(*
SPDX-FileCopyrightText: © 2026 Oleksandr Tiutyk <trofimich@gmail.com>
SPDX-License-Identifier: MIT
License: https://opensource.org/license/mit
*)

(*!
<summary>Enumerates allocated text fragments from a borrowed source string.</summary>
<description>
Initialization requires a separator containing 1 to 80 characters, stored in a fixed buffer. The source must
remain alive and unchanged during iteration. The enumerator owns the current fragment; borrowed fragment
references expire on MoveNext, Reset or destruction. Allocation failure uses the terminal memory mechanism.
With a nonempty separator, empty fragments are preserved when RemoveEmptyEntries is FALSE, including the final
fragment after a trailing separator and one fragment for an empty source. RemoveEmptyEntries filters empty
fragments after optional trimming. MaxCount still limits the number of returned fragments. Do not copy an
instance by assignment or pass it by value while it owns an allocated buffer; use references instead.
Assignment does not clone the buffer or transfer ownership. Do not overwrite an instance that still owns a
buffer. The creator is responsible for the splitter lifetime and cleanup. Release the current fragment with
Reset when abandoning iteration. Delete the splitter itself only if it was allocated with __NEW; FB_exit
releases its current fragment. Statically or locally declared instances must not be passed to __DELETE. The
borrowed source is never owned or freed by the splitter.
</description>
*)

{attribute 'no_explicit_call' := 'do not call this function block directly'}
FUNCTION_BLOCK WideStringSplittingEnumerator EXTENDS Object IMPLEMENTS IEnumerator
VAR_OUTPUT
	SourceString : POINTER TO WSTRING;
	SourceStringLength : UDINT;
	SourceStringSize : UDINT;
	Separator : WSTRING(80);
	SeparatorLength : UDINT;
	//!<summary>
	//! Maximum number of returned fragments; zero means unlimited. Empty fragments removed after optional
	//! trimming do not count toward the limit. Remaining text is not returned after the limit is reached and is
	//! not merged into the last fragment.
	//! </summary>
	MaxCount : UDINT := 0;
	TrimEntries : BOOL := FALSE;
	RemoveEmptyEntries : BOOL := FALSE;	
END_VAR
VAR_STAT
	//! <summary>Class name shared by all instances of this function block.</summary>
	{attribute 'hide'} 
	_ClassName : STRING := __POUNAME();
END_VAR
VAR
	{attribute 'hide'} 
	_CurrentString : POINTER TO WSTRING;
	{attribute 'hide'} 
	_CurrentStringLength : UDINT;
	{attribute 'hide'} 
	_CurrentEntry : POINTER TO WSTRING;
	{attribute 'hide'} 
	_CurrentEntrySize : UDINT;
	{attribute 'hide'} 
	_EntryCount : UDINT; 
END_VAR

{attribute 'monitoring' := 'call'}
PROPERTY ClassName : REFERENCE TO STRING
GET
ClassName REF= _ClassName;
END_GET
END_PROPERTY

(*!
<summary>Returns a borrowed generic view of the current split fragment.</summary>
<description>
The descriptor does not own the fragment. With no current fragment it is reset to a null generic value. The
descriptor is reused by this getter; do not modify it or retain its payload across MoveNext, Reset or
destruction. Copy the text for independent storage. Descendants cannot override this cursor operation;
advancement, reset and borrowed current views use the same cursor state.
</description>
*)

{attribute 'monitoring' := 'call'}
PROPERTY FINAL Current : REFERENCE TO GENERIC_VALUE
GET
VAR_INST
	genericValue : GENERIC_VALUE;
END_VAR
IF _CurrentEntry <> 0 AND_THEN _CurrentEntrySize > 0 THEN
	genericValue := GenericValueFactory.FromParts(
		genericTypeClass := GENERIC_TYPE_CLASS.STRING_16,
		address := _CurrentEntry,
		size := _CurrentEntrySize,
		memoryManagementBehavior := GENERIC_MEMORY_MANAGEMENT_BEHAVIOR.STORE_ORIGINAL_REFERENCE_AND_NOT_OWNS_MEMORY
	);
ELSE
	genericValue.Reset();
END_IF

Current REF= genericValue;
END_GET
END_PROPERTY

(*!
<summary>Returns a borrowed reference to the current split fragment.</summary>
<description>
The reference is invalid when no current fragment exists. Do not retain it across MoveNext, Reset or
destruction; copy the text if it must outlive cursor advancement. Descendants cannot override this cursor
operation; advancement, reset and borrowed current views use the same cursor state.
</description>
*)
PROPERTY FINAL CurrentEntry : REFERENCE TO WSTRING
GET
IF _CurrentEntry <> 0 THEN
	CurrentEntry REF= _CurrentEntry^;	
END_IF
END_GET
END_PROPERTY

(*!
<summary>Releases the cursor-owned fragment buffer.</summary>
<description>
Does not release the borrowed source string. Destruction invalidates references to the current fragment and
must not raise exceptions.
</description>
*)
//!<param name="bInCopyCode">
//! if TRUE, the exit method is called for exiting an instance that is copied afterwards (online change).
//! </param>

METHOD FB_exit : BOOL
VAR_INPUT
	
	bInCopyCode	: BOOL;
END_VAR
IF _CurrentEntry <> 0 THEN
	__DELETE(_CurrentEntry);
END_IF
END_METHOD

(*!
<summary>Sets the borrowed source and splitting options, then resets iteration.</summary>
<description>
SourceStringLength counts UTF-16 code units; SourceStringSize counts bytes including the terminator. The
separator is copied into internal storage. The source remains caller-owned. Descendants cannot override this
cursor operation; advancement, reset and borrowed current views use the same cursor state.
</description>
*)
//!<param name="maxCount">
//! Maximum number of returned fragments; zero means unlimited. Empty fragments removed after optional
//! trimming do not count toward the limit. Remaining text is not returned after the limit is reached and is
//! not merged into the last fragment.
//! </param>
//!<param name="separator">
//! Separator containing 1 to 80 characters; the caller must validate its length before initialization.
//! </param>
METHOD INTERNAL FINAL Initialize
VAR_INPUT
	sourceString : POINTER TO WSTRING;
	separator : WSTRING(80);
	maxCount : UDINT;
	trimEntries : BOOL;
	removeEmptyEntries : BOOL;
END_VAR
THIS^.SourceString := sourceString;
THIS^.SourceStringLength := WideStrings.InternalGetLength(value := sourceString);
THIS^.SourceStringSize := (THIS^.SourceStringLength + 1) * WideStrings.CharSize; 
THIS^.Separator := separator;
THIS^.SeparatorLength := WideStrings.InternalGetLength(value := ADR(THIS^.Separator));
THIS^.MaxCount := maxCount;
THIS^.TrimEntries := trimEntries;
THIS^.RemoveEmptyEntries := removeEmptyEntries;

_CurrentString := THIS^.SourceString;

Reset();
END_METHOD

(*!
<summary>Releases the previous fragment and advances to the next selected fragment.</summary>
<description>
Returns TRUE when a new current fragment is available, FALSE at the end or when the configured limit is
reached. A non-null cursor with zero remaining length represents a pending empty final fragment; a null cursor
marks completed iteration. Empty fragments are returned unless RemoveEmptyEntries is TRUE, subject to
MaxCount. Each fragment owns a null-terminated allocation; allocation failure invokes
DynamicMemoryManager.RaiseAllocationFailure before the buffer is accessed. Descendants cannot override this
cursor operation; advancement, reset and borrowed current views use the same cursor state.
</description>
*)
METHOD FINAL MoveNext : BOOL
VAR
	separatorPosition : UDINT;
END_VAR
START:

IF _CurrentEntry <> 0 THEN
	_CurrentEntrySize := 0;
	
	__DELETE(_CurrentEntry);
END_IF

IF _CurrentString = 0 OR_ELSE Separator = "" OR_ELSE (MaxCount > 0 AND_THEN _EntryCount >= MaxCount) THEN
	RETURN;
END_IF

IF WideStrings.InternalFind(
	stringToSearchIn := _CurrentString,
	stringToSearchInLength := _CurrentStringLength,
	stringToFind := ADR(Separator),
	stringToFindLength := SeparatorLength,
	position => separatorPosition
) THEN
	_CurrentEntrySize := separatorPosition * WideStrings.CharSize;
	_CurrentEntry := __NEW(BYTE, _CurrentEntrySize);

	IF _CurrentEntry = 0 THEN
		DynamicMemoryManager.RaiseAllocationFailure();
	END_IF

	Tc2_System.MEMCPY(
		destAddr := _CurrentEntry,
		srcAddr := _CurrentString,
		n := (separatorPosition - 1) * WideStrings.CharSize
	);
	Tc2_System.MEMSET(
		destAddr := _CurrentEntry + ((separatorPosition - 1) * WideStrings.CharSize),
		fillByte := 0,
		n := WideStrings.CharSize
	);

	_CurrentString := _CurrentString + ((separatorPosition - 1) * WideStrings.CharSize) + (SeparatorLength * WideStrings.CharSize);
	_CurrentStringLength := _CurrentStringLength - separatorPosition + 1 - SeparatorLength;
ELSE	
	_CurrentEntrySize := (_CurrentStringLength + 1) * WideStrings.CharSize;	
	_CurrentEntry := __NEW(BYTE, _CurrentEntrySize);

	IF _CurrentEntry = 0 THEN
		DynamicMemoryManager.RaiseAllocationFailure();
	END_IF
	
	Tc2_System.MEMCPY(destAddr := _CurrentEntry, srcAddr := _CurrentString, n := _CurrentEntrySize);
	
	_CurrentString := 0;
	_CurrentStringLength := 0;
END_IF

IF TrimEntries THEN
	WideStrings.TrimChar(stringToTrim := _CurrentEntry^);
END_IF

IF RemoveEmptyEntries AND_THEN _CurrentEntry^ = "" THEN
	JMP START;
END_IF

_EntryCount := _EntryCount + 1;

MoveNext := TRUE;
END_METHOD

(*!
<summary>Provides the library namespace used in diagnostics.</summary>
<description>
Borrowed read-only reference to the compiler-initialized library namespace; no ownership transfer.
</description>
*)
{attribute 'monitoring' := 'call'}
PROPERTY NamespaceName : REFERENCE TO STRING
GET
NamespaceName REF= CurrentNamespace.Name;
END_GET
END_PROPERTY

(*!
<summary>Releases the current fragment and resets iteration to before the first entry.</summary>
<description>
Preserves splitting settings and does not allocate memory or modify the source string. Previously borrowed
fragment addresses and references become invalid. The initialized source string must remain alive and
unchanged throughout iteration. Repeated Reset calls are allowed, including before iteration and after its
end. Descendants cannot override this cursor operation; advancement, reset and borrowed current views use the
same cursor state.
</description>
*)
METHOD FINAL Reset
IF _CurrentEntry <> 0 THEN
	__DELETE(_CurrentEntry);
END_IF

_CurrentEntry := 0;
_CurrentEntrySize := 0;

_CurrentString := SourceString;
_CurrentStringLength := SourceStringLength;
_EntryCount := 0;
END_METHOD

(*!
<summary>Reports the byte size of this concrete instance.</summary>
<description>
Uses XSIZEOF on the instance. Does not include separately allocated payloads or prove that an arbitrary
address is valid.
</description>
*)
{attribute 'monitoring' := 'call'}
PROPERTY SelfSize : ULINT
GET
SelfSize := XSIZEOF(THIS^);
END_GET
END_PROPERTY

END_FUNCTION_BLOCK

(* stored: Version 1.1.0.1
   POU WideStringSplittingEnumerator: Id {cd3c3f30-cd38-4659-b9c4-859e877b4baf}, SpecialFunc None
   Property ClassName: Id {eb782797-fea3-47ac-a8db-cbfc72d737be}
   Get Get: Id {b0de37f0-477e-4092-a2e4-1e3cd48b7e08}
   Property Current: Id {a33a22ac-5669-4623-936f-19fdd6a797a9}
   Get Get: Id {b343fd78-0841-4c7a-bd2d-6b447815e0a9}
   Property CurrentEntry: Id {f4b2ce05-56f1-4a2a-ab8a-2d63ad7de743}
   Get Get: Id {859e54d6-429d-47fd-a753-3e8e965a0bc3}
   Method FB_exit: Id {d23faa7c-5379-472c-b75f-ff9aa468fe1d}
   Method Initialize: Id {efd8c83e-84af-4552-92cf-49864ca5b37a}
   Method MoveNext: Id {6f4c66bb-70e6-443d-b741-5ac7aedc0a0c}
   Property NamespaceName: Id {606a15c2-aeca-432d-8e3c-a9852072d07e}
   Get Get: Id {8d26a153-dac4-4ce7-b323-94027a2445d2}
   Method Reset: Id {6ff5f895-f51d-4f1c-b79b-00ce34e370cc}
   Property SelfSize: Id {e6e7cb18-6bbe-4fa5-8b86-e60c4005ed50}
   Get Get: Id {6cd74453-76de-45a9-9aff-7d3ec88a250f} *)
